Fanuc KAREL source: KA00176.KL

PROGRAM KA00176
%NOLOCKGROUP
VAR
  SRC: ARRAY[4] OF STRING[20]
  DST: ARRAY[4] OF BYTE
BEGIN
  DST = SRC
END KA00176
